(* IEC 61131-3 sources: ZPLC/conformance/rt, 6 files *)

(* ---- rt-006-runaway-loop-ends-in-a-fault.st ---- *)
PROGRAM Runaway
VAR
  count AT %QW0 : INT;
END_VAR
  WHILE TRUE DO
    count := count + 1;
  END_WHILE;
END_PROGRAM

(* ---- rt-007-vm-fault-drives-outputs-safe.st ---- *)
PROGRAM Safe
VAR
  zero : INT;
  lamp AT %QX0.0 : BOOL;
  other AT %QW1 : INT;
END_VAR
  lamp := TRUE;
  other := 100 / zero;
END_PROGRAM

(* ---- rt-015-event-triggered-task-is-rejected.st ---- *)
PROGRAM OnEvent
VAR
  runs AT %QW0 : INT;
END_VAR
  runs := runs + 1;
END_PROGRAM

(* ---- rt-015-two-cyclic-tasks-with-different-intervals-slow.st ---- *)
PROGRAM Slow
VAR
  runs AT %QW1 : INT;
END_VAR
  runs := runs + 1;
END_PROGRAM

(* ---- rt-015-two-cyclic-tasks-with-different-intervals.st ---- *)
PROGRAM Fast
VAR
  runs AT %QW0 : INT;
END_VAR
  runs := runs + 1;
END_PROGRAM

(* ---- rt-034-watchdog-reset-is-reported-and-changes-nothing.st ---- *)
PROGRAM Feed
VAR
  before AT %QW0 : INT;
  after AT %QW1 : INT;
  scans AT %QW2 : INT;
END_VAR
  before := 7;
  WATCHDOG_RESET();
  after := before + 1;
  scans := scans + 1;
END_PROGRAM
